// TIA Portal V19 export
DATA_BLOCK "MOTOR_DB"   // DB24
// stored: InstanceOfName MOTOR, InstanceOfType FB
"MOTOR"
   // VAR
   //    AG_01 { S7_SetPoint := 'True'} : "MOTOR_FB1";
   // END_VAR
BEGIN
END_DATA_BLOCK
